(* PLC project zarechnaya.project, CODESYS CODESYS V3.5 SP17 Patch 3 *)
(* stored: creationDateTime 2026-10-20T05:42:22.1976194, modificationDateTime 1601-01-01T03:00:00 *)

(* FB_LevelAlarm — сигнализация уровня в фильтре (FBD, 4 сети, Jump/Label). Поведение (модель scenarios/reference/model_FB_LevelAlarm.py): 1. xHigh := rLevel > rHigh; 2. если NOT xEnable — переход на lblOut (сеть 3 пропускается, тревога держит прошлое значение); 3. xAlarm := (xHigh OR xAlarm) AND NOT xAck — защёлка с квитированием; 4. (метка lblOut) xLamp := xAlarm AND xEnable. *)
FUNCTION_BLOCK FB_LevelAlarm
  VAR_INPUT
    rLevel : REAL;
    rHigh : REAL;
    xEnable : BOOL;
    xAck : BOOL;
  END_VAR
  VAR_OUTPUT
    xAlarm : BOOL;
    xLamp : BOOL;
  END_VAR
  VAR
    xHigh : BOOL;
  END_VAR

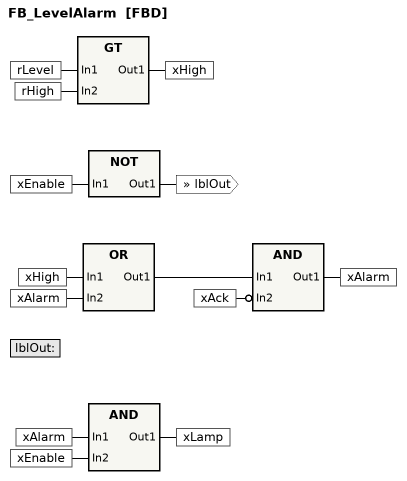
(* FBD diagram, written out as Structured Text *)
xHigh := rLevel > rHigh;
(* --- network: Пропуск при выводе из работы --- *)
IF NOT xEnable THEN JMP lblOut; END_IF;
(* --- network: Защёлка тревоги --- *)
xAlarm := (xHigh OR xAlarm) AND NOT xAck;
lblOut:
(* --- network: Лампа --- *)
xLamp := xAlarm AND xEnable;
END_FUNCTION_BLOCK
